Universal Robots PolyScope program: Retract.urp

Program Retract (createdIn=3.0.0 lastSavedIn=3.0.0 directory=/programs installation=default)
Robot Program (runOnlyOnce=true motionType=MoveJ speed=1.047198 acceleration=1.396263 useActiveTCP=false)
  'Program generated by VerticalBot Studio for UR10 on 25/10/2026 12:00:00'
  'Using nominal kinematics.'
  'Using Ref. Frame 2: p[-0.800000, 0.500000, 0.100000, 0.000000, 0.000000, 3.141593]'
  'Using TCP Paint gun: p[0.050000, 0.000000, 0.450000, 0.000000, 0.523599, 0.000000]'
  Script: set_tcp(p[0.050000, 0.000000, 0.450000, 0.000000, 0.523599, 0.000000])
  MoveL speed 250 mm/s, acceleration 1200 mm/s^2 (useActiveTCP=true)
    Waypoint Waypoint_1: TCP in base x=-825.987 y=133.387 z=269.825 mm, rx=-2.6833 ry=0.2664 rz=0.0605 rad; joints [-153.215, -81.897, -104.364, -66.506, 50.655, 115.012] deg; flange x=-647.838 y=-77.959 z=628.428 mm, rx=-2.5528 ry=0.0987 rz=0.7461 rad
  Script: movej([-2.652656, -1.365240, -1.512183, -1.127521, 1.275171, 1.920421],1.20000,0.75000,0,0.0000)
  MoveJ speed 42.97 deg/s, acceleration 68.75 deg/s^2 (useActiveTCP=true)
    Waypoint Waypoint_2: TCP in base x=-866.761 y=-115.117 z=513.712 mm, rx=3.1014 ry=0.052 rz=-0.3627 rad; joints [-151.986, -78.222, -86.642, -64.602, 73.062, 110.032] deg; flange x=-594.55 y=-100.237 z=875.208 mm, rx=2.8946 ry=0.0426 rz=-1.1501 rad
